TYPE U_LintUnion :
UNION
    nDword : DWORD;
    arBytes : ARRAY[0..3] OF BYTE;
END_UNION
END_TYPE

(* stored: Version 1.1.0.1, ProductVersion 3.1.4026.18
   DUT U_LintUnion: Id {c547fb77-8233-03e5-043a-2c4f51bc998e} *)
